// TIA Portal V19 export
DATA_BLOCK "RUA_R4_DB"   // DB45
// stored: InstanceOfName RUA_R4, InstanceOfType FB
"RUA_R4"
   // VAR
   //    START_Instance { S7_SetPoint := 'True'} : "START";
   //    "HEAT/COOL_Instance" { S7_SetPoint := 'True'} : "HEAT/COOL";
   //    "AUTO_COOLING_UTIITY SELECTION_Instance" { S7_SetPoint := 'True'} : "AUTO_COOLING_UTIITY SELECTION";
   //    AUTO_HEATING_SELECTION_Instance { S7_SetPoint := 'True'} : "AUTO_HEATING_SELECTION";
   //    "SEMI/_AUTO_Instance" { S7_SetPoint := 'True'} : "SEMI/_AUTO";
   //    COOLING_PROCESS_Instance { S7_SetPoint := 'True'} : "COOLING_PROCESS";
   //    HEATING_PROCEES_Instance { S7_SetPoint := 'True'} : "HEATING_PROCEES";
   //    RAMP_Instance { S7_SetPoint := 'True'} : "RAMP";
   // END_VAR
BEGIN
END_DATA_BLOCK
